Fanuc KAREL source: kd00065.KL

-- PROVISIONAL review KL for V1013-1; original PC SHA256 caa4a0f15524ce1b17b1828e34a062e2bb7aa46a94f5e5b599fde58edbe714e6
-- Incomplete behavior may be omitted. Consult companion uncertainty JSON. Do not deploy.
PROGRAM KD00065
%NOLOCKGROUP
VAR
  I : INTEGER
  J : INTEGER
  B : BOOLEAN
  R : REAL
  S : STRING[80]
BEGIN
  -- UNRESOLVED_PC offsets 5-17; opcodes 9D,81,18,9D,1B,9D,12,13,04
  -- UNRESOLVED_PC offsets 22-26; opcodes 7F
END KD00065
